(* Logix 5000 project; controller SmartManufacturingCell Emulate 5570 rev 33.11; software revision 33.03; part 2 of 5 *)
(* tags used below, declared in another part *)
   ExitDischargeTimeout : TIMER;   // Non-retentive timer; preset in milliseconds.
   ExitResetONS : BOOL;
   Inspection_RejectSample : BOOL;
   Inspection_StateAtScan : DINT;
   InspectionProcessDelay : TIMER;   // Non-retentive timer; preset in milliseconds.
   InspectionResetONS : BOOL;
   InspectionTimeout : TIMER;   // Non-retentive timer; preset in milliseconds.
   Reject_AutoExtendAllowed : BOOL;
   Reject_ManualExtendAllowed : BOOL;
   Reject_ManualExtendArmed : BOOL;
   Reject_ResetAllowed : BOOL;   // Reject recovery conditions satisfied; permits a fresh Reset request.
   RejectExtendTimeout : TIMER;   // Non-retentive timer; preset in milliseconds.
   RejectResetONS : BOOL;
   RejectRetractTimeout : TIMER;   // Non-retentive timer; preset in milliseconds.
   Cfg_InspectionTimeMs : DINT;   // Inspection duration; 100..2000 ms. Sampled when inspection starts.
   Exit_Flt_DischargeTimeout : BOOL;   // Good or reject bottle departure not confirmed within 3 s Latched; clear cell, remove cause, then fresh Reset.
   Exit_Sts_ResetAccepted : BOOL;   // Exit Sts ResetAccepted
   Exit_Sts_State : DINT;   // 0 Empty; 10 Waiting; 20 Good discharge; 30 Extending; 40 Reject discharge; 50 Retracting; 60 Complete; 90 Faulted
   HMI_Cmd_ClearCell : BOOL;   // Request removal of simulated bottles during fault recovery
   HMI_Cmd_LoadBottle : BOOL;   // Request one simulated bottle at the available entry position
   HMI_Cmd_RejectExtend : BOOL;
   HMI_Cmd_Reset : BOOL;   // Request fault reset after recovery conditions are satisfied
   HMI_Cmd_Stop : BOOL;   // Request controlled production stop
   HMI_Sim_InspectionFailToComplete : BOOL;   // Prevent inspection process timer from completing. Simulation test only.
   HMI_Sim_NextInspectionRejects : BOOL;   // Select Reject for the next inspection
   Inspection_Flt_Timeout : BOOL;   // Inspection did not finish within 3 s Latched; clear cell, remove cause, then fresh Reset.
   Inspection_Sts_ResetAccepted : BOOL;   // Inspection Sts ResetAccepted
   Inspection_Sts_State : DINT;   // 0 Empty; 10 Waiting; 20 Inspecting; 40 Complete; 90 Faulted
   Production_Bottles : UDT_Bottle[4];
   Production_Sts_ClearCellAccepted : BOOL;
   Production_Sts_LoadAccepted : BOOL;
   Production_Sts_LoadAllowed : BOOL;
   Production_Sts_LoadBlockReason : DINT;   // 0 allowed; 10 not Auto Running/ProcessStations; 20 command conflict; 30 conveyor moving; 40 Entry occupied; 50 fault/sta
   Production_Sts_SequenceState : DINT;   // 0 = Idle 10 = ProcessStations 20 = Indexing 30 = ConfirmPositions
   Reject_Flt_FailToExtend : BOOL;   // Reject actuator did not extend within 2 s Latched; clear cell, remove cause, then fresh Reset.
   Reject_Flt_FailToRetract : BOOL;   // Reject actuator did not retract within 2 s Latched; clear cell, remove cause, then fresh Reset.
   Reject_Sts_BlockReason : DINT;   // Reason manual reject extension is unavailable. 0 = Ready to accept Extend. 10 = Release Extend to rearm. 20 = Good-bottl
   Reject_Sts_ResetAccepted : BOOL;
   Sim_In_ConveyorRunning : BOOL;   // Simulated conveyor movement feedback
   Sim_In_EntryPE : BOOL;   // Simulated bottle detected at entry
   Sim_In_GoodExitPE : BOOL;   // Bottle detected passing through good discharge path
   Sim_In_InspectionPE : BOOL;   // Simulated bottle detected at inspection position
   Sim_In_RejectExitPE : BOOL;   // Bottle detected passing through reject discharge path
   Sim_In_RejectExtended : BOOL;   // Simulated reject actuator confirmed extended
   Sim_In_RejectRetracted : BOOL;   // Simulated reject actuator confirmed retracted
   Sim_Out_ConveyorRun : BOOL;   // Command simulated conveyor to run
   Sim_Out_GoodDischargeRun : BOOL;   // Command simulated good-bottle discharge mechanism to run
   Sim_Out_RejectExtend : BOOL;   // Command simulated reject actuator to extend
   Sys_Sts_AutoMode : BOOL;   // Auto mode accepted and active
   Sys_Sts_BlockingFault : BOOL;   // Active blocking fault prevents production and manual equipment operation.
   Sys_Sts_MachineState : DINT;   // 0 = Stopped 10 = Running 20 = Stopping 30 = Faulted
   Sys_Sts_ManualMode : BOOL;   // Manual mode accepted and active
   Sys_Sts_ResetAllowed : BOOL;   // Sys Sts ResetAllowed
   Sys_Sts_StartupReady : BOOL;   // Sys Sts StartupReady
(* Program_Inspection, continued *)

ROUTINE Exit_Faults   (* ladder *)
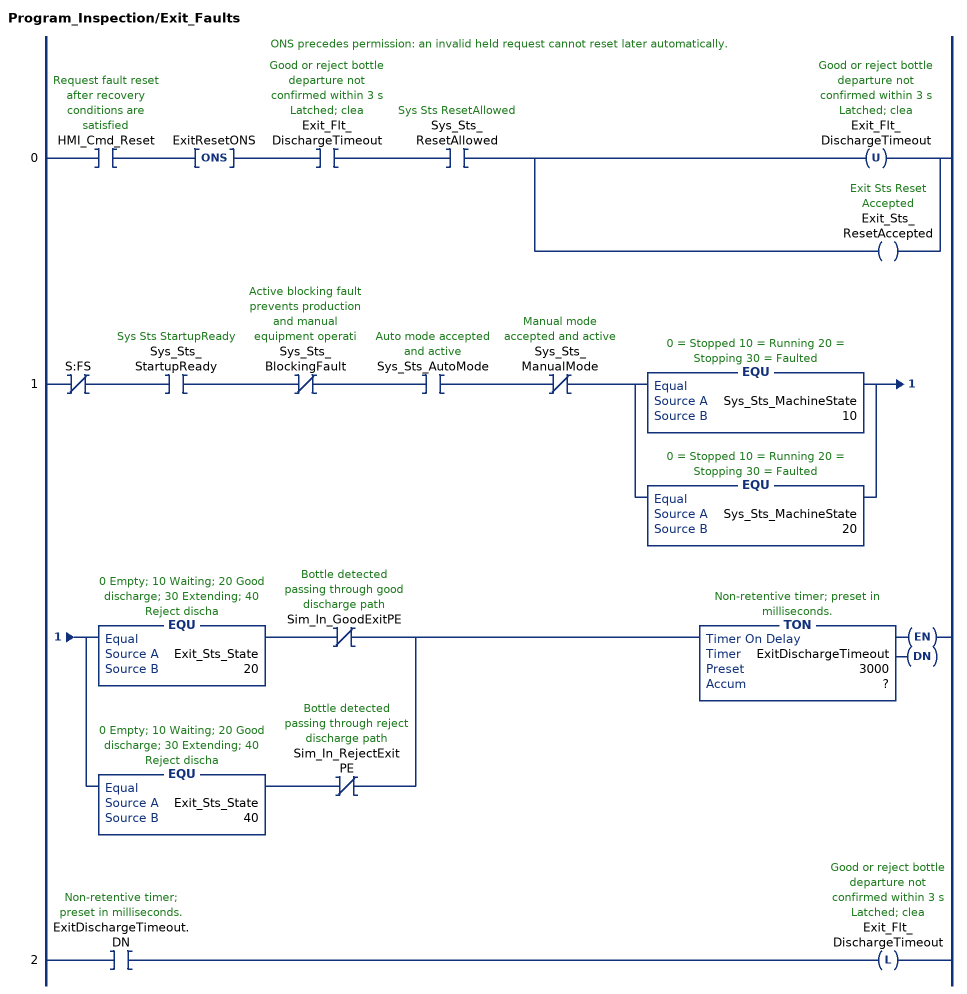
   // ONS precedes permission: an invalid held request cannot reset later automatically.
   0: XIC(HMI_Cmd_Reset)ONS(ExitResetONS)XIC(Exit_Flt_DischargeTimeout)XIC(Sys_Sts_ResetAllowed)[OTU(Exit_Flt_DischargeTimeout) ,OTE(Exit_Sts_ResetAccepted) ];
   1: XIO(S:FS)XIC(Sys_Sts_StartupReady)XIO(Sys_Sts_BlockingFault)XIC(Sys_Sts_AutoMode)XIO(Sys_Sts_ManualMode)[EQU(Sys_Sts_MachineState,10) ,EQU(Sys_Sts_MachineState,20) ][EQU(Exit_Sts_State,20) XIO(Sim_In_GoodExitPE) ,EQU(Exit_Sts_State,40) XIO(Sim_In_RejectExitPE) ]TON(ExitDischargeTimeout,?,?);
   2: XIC(ExitDischargeTimeout.DN)OTL(Exit_Flt_DischargeTimeout);
END_ROUTINE

ROUTINE Inspection_Control   (* ladder *)
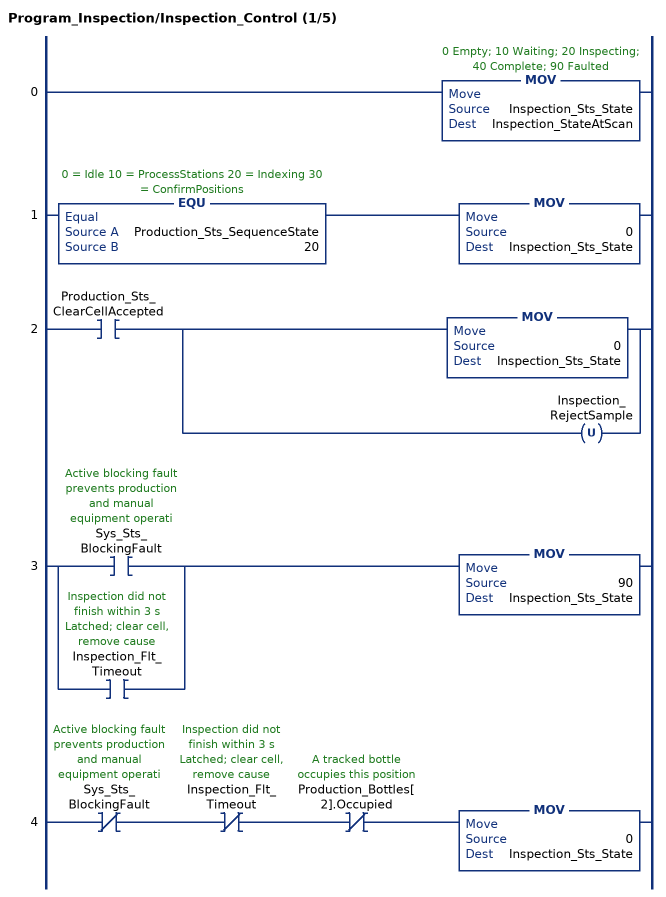
   0: MOV(Inspection_Sts_State,Inspection_StateAtScan);
   1: EQU(Production_Sts_SequenceState,20)MOV(0,Inspection_Sts_State);
   2: XIC(Production_Sts_ClearCellAccepted)[MOV(0,Inspection_Sts_State) ,OTU(Inspection_RejectSample) ];
   3: [XIC(Sys_Sts_BlockingFault) ,XIC(Inspection_Flt_Timeout) ]MOV(90,Inspection_Sts_State);
   4: XIO(Sys_Sts_BlockingFault)XIO(Inspection_Flt_Timeout)XIO(Production_Bottles[2].Occupied)MOV(0,Inspection_Sts_State);
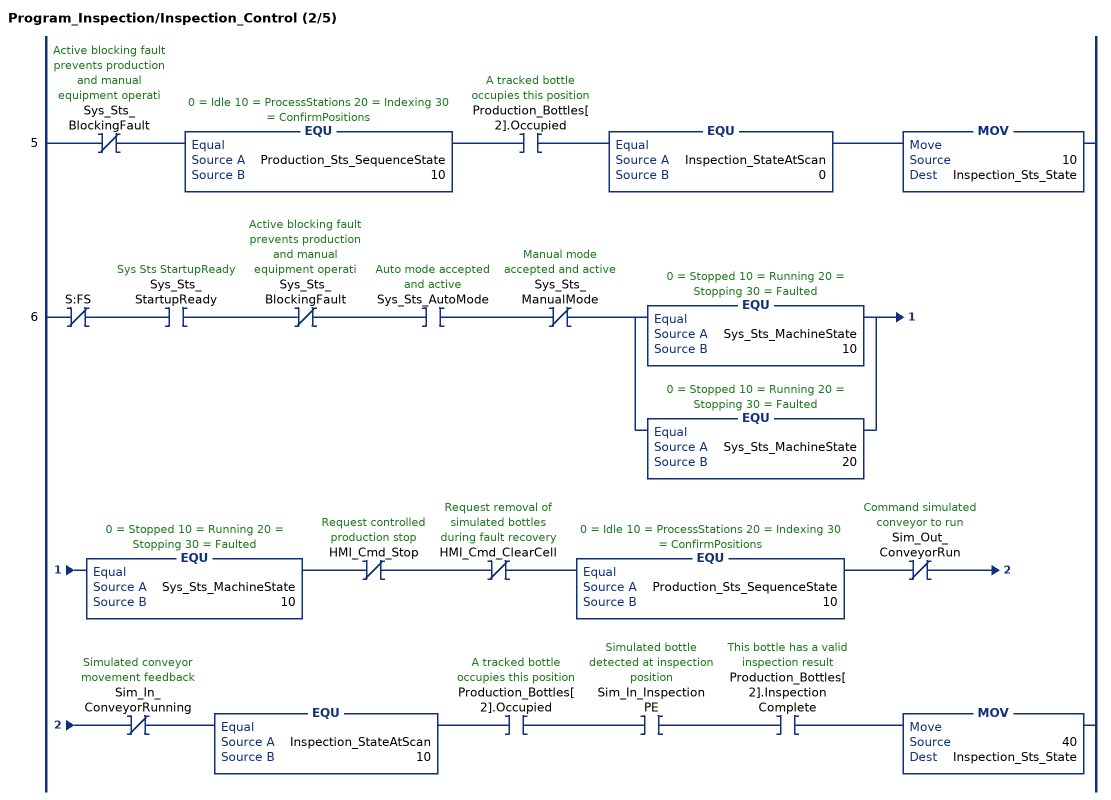
   5: XIO(Sys_Sts_BlockingFault)EQU(Production_Sts_SequenceState,10)XIC(Production_Bottles[2].Occupied)EQU(Inspection_StateAtScan,0)MOV(10,Inspection_Sts_State);
   6: XIO(S:FS)XIC(Sys_Sts_StartupReady)XIO(Sys_Sts_BlockingFault)XIC(Sys_Sts_AutoMode)XIO(Sys_Sts_ManualMode)[EQU(Sys_Sts_MachineState,10) ,EQU(Sys_Sts_MachineState,20) ]EQU(Sys_Sts_MachineState,10)XIO(HMI_Cmd_Stop)XIO(HMI_Cmd_ClearCell)EQU(Production_Sts_SequenceState,10)XIO(Sim_Out_ConveyorRun)XIO(Sim_In_ConveyorRunning)EQU(Inspection_StateAtScan,10)XIC(Production_Bottles[2].Occupied)XIC(Sim_In_InspectionPE)XIC(Production_Bottles[2].InspectionComplete)MOV(40,Inspection_Sts_State);
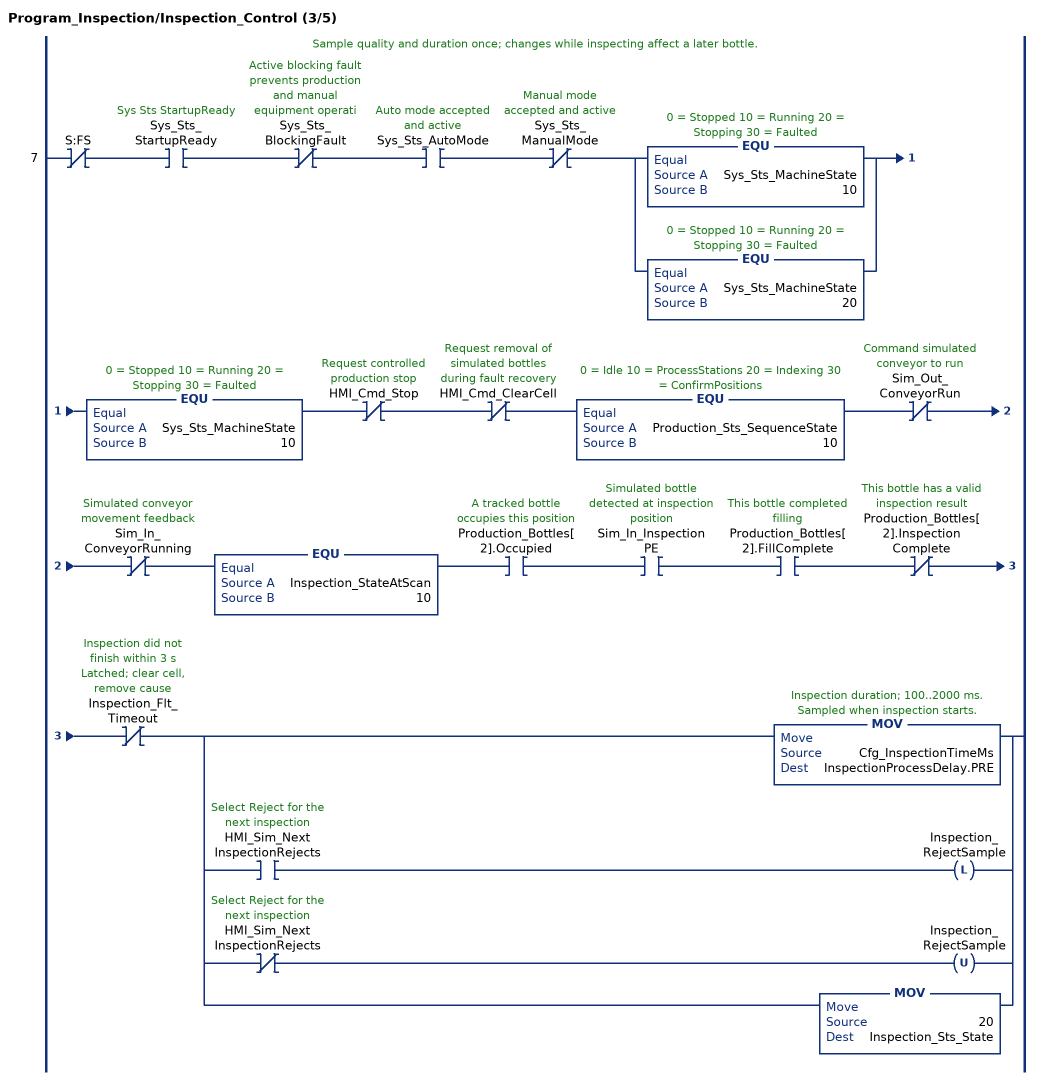
   // Sample quality and duration once; changes while inspecting affect a later bottle.
   7: XIO(S:FS)XIC(Sys_Sts_StartupReady)XIO(Sys_Sts_BlockingFault)XIC(Sys_Sts_AutoMode)XIO(Sys_Sts_ManualMode)[EQU(Sys_Sts_MachineState,10) ,EQU(Sys_Sts_MachineState,20) ]EQU(Sys_Sts_MachineState,10)XIO(HMI_Cmd_Stop)XIO(HMI_Cmd_ClearCell)EQU(Production_Sts_SequenceState,10)XIO(Sim_Out_ConveyorRun)XIO(Sim_In_ConveyorRunning)EQU(Inspection_StateAtScan,10)XIC(Production_Bottles[2].Occupied)XIC(Sim_In_InspectionPE)XIC(Production_Bottles[2].FillComplete)XIO(Production_Bottles[2].InspectionComplete)XIO(Inspection_Flt_Timeout)[MOV(Cfg_InspectionTimeMs,InspectionProcessDelay.PRE) ,XIC(HMI_Sim_NextInspectionRejects) OTL(Inspection_RejectSample) ,XIO(HMI_Sim_NextInspectionRejects) OTU(Inspection_RejectSample) ,MOV(20,Inspection_Sts_State) ];
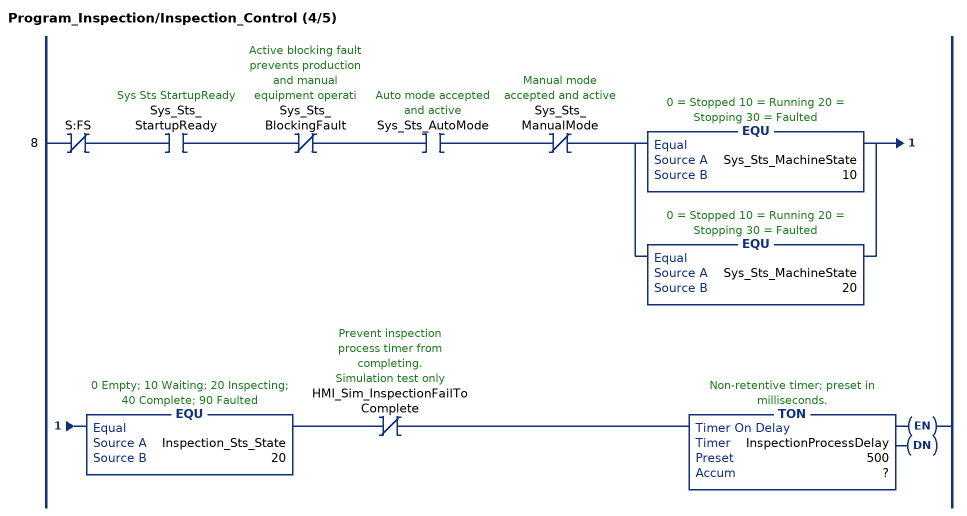
   8: XIO(S:FS)XIC(Sys_Sts_StartupReady)XIO(Sys_Sts_BlockingFault)XIC(Sys_Sts_AutoMode)XIO(Sys_Sts_ManualMode)[EQU(Sys_Sts_MachineState,10) ,EQU(Sys_Sts_MachineState,20) ]EQU(Inspection_Sts_State,20)XIO(HMI_Sim_InspectionFailToComplete)TON(InspectionProcessDelay,?,?);
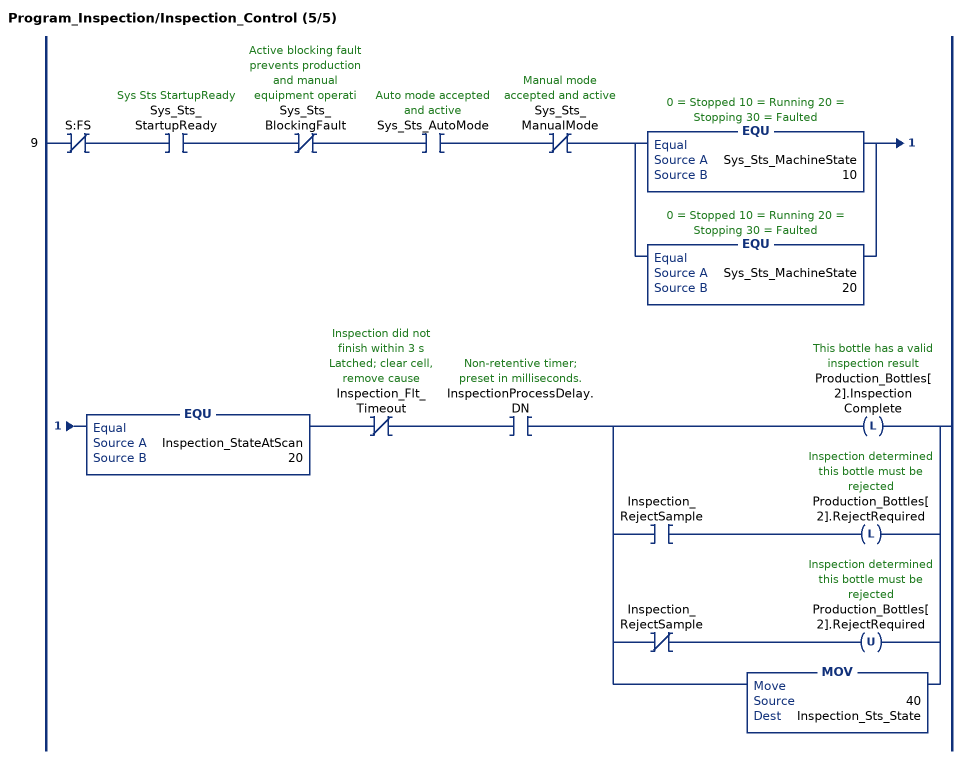
   9: XIO(S:FS)XIC(Sys_Sts_StartupReady)XIO(Sys_Sts_BlockingFault)XIC(Sys_Sts_AutoMode)XIO(Sys_Sts_ManualMode)[EQU(Sys_Sts_MachineState,10) ,EQU(Sys_Sts_MachineState,20) ]EQU(Inspection_StateAtScan,20)XIO(Inspection_Flt_Timeout)XIC(InspectionProcessDelay.DN)[OTL(Production_Bottles[2].InspectionComplete) ,XIC(Inspection_RejectSample) OTL(Production_Bottles[2].RejectRequired) ,XIO(Inspection_RejectSample) OTU(Production_Bottles[2].RejectRequired) ,MOV(40,Inspection_Sts_State) ];
END_ROUTINE

ROUTINE Inspection_Faults   (* ladder *)
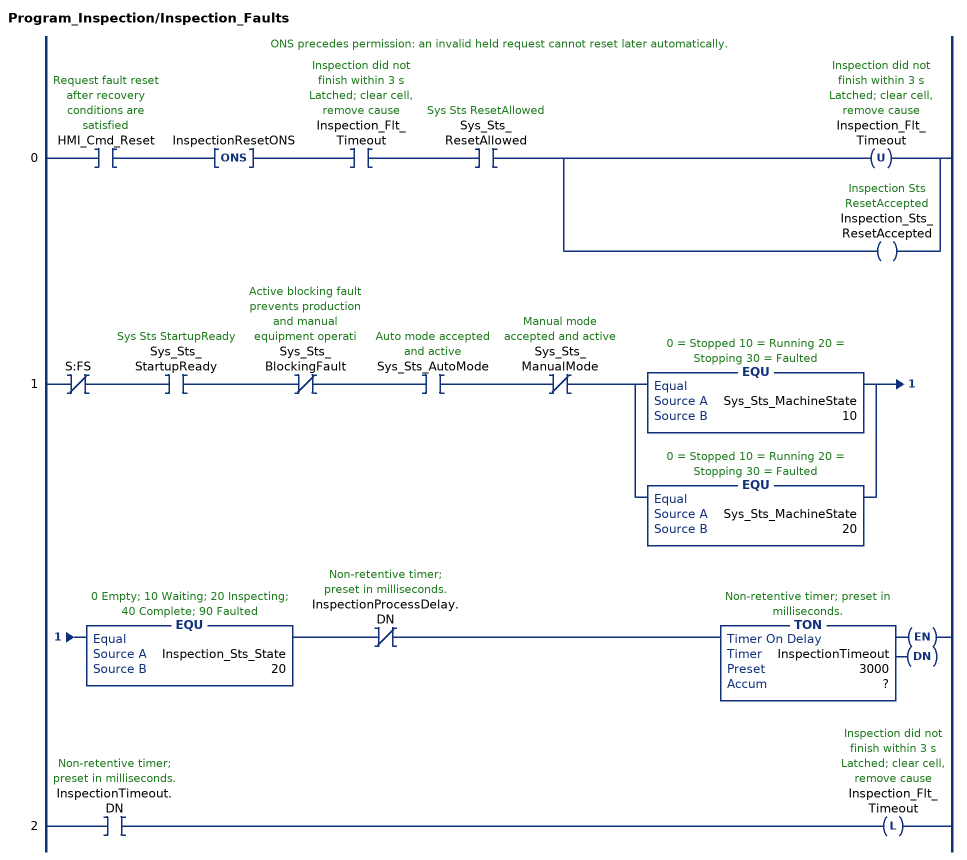
   // ONS precedes permission: an invalid held request cannot reset later automatically.
   0: XIC(HMI_Cmd_Reset)ONS(InspectionResetONS)XIC(Inspection_Flt_Timeout)XIC(Sys_Sts_ResetAllowed)[OTU(Inspection_Flt_Timeout) ,OTE(Inspection_Sts_ResetAccepted) ];
   1: XIO(S:FS)XIC(Sys_Sts_StartupReady)XIO(Sys_Sts_BlockingFault)XIC(Sys_Sts_AutoMode)XIO(Sys_Sts_ManualMode)[EQU(Sys_Sts_MachineState,10) ,EQU(Sys_Sts_MachineState,20) ]EQU(Inspection_Sts_State,20)XIO(InspectionProcessDelay.DN)TON(InspectionTimeout,?,?);
   2: XIC(InspectionTimeout.DN)OTL(Inspection_Flt_Timeout);
END_ROUTINE

ROUTINE MainRoutine   (* ladder *)
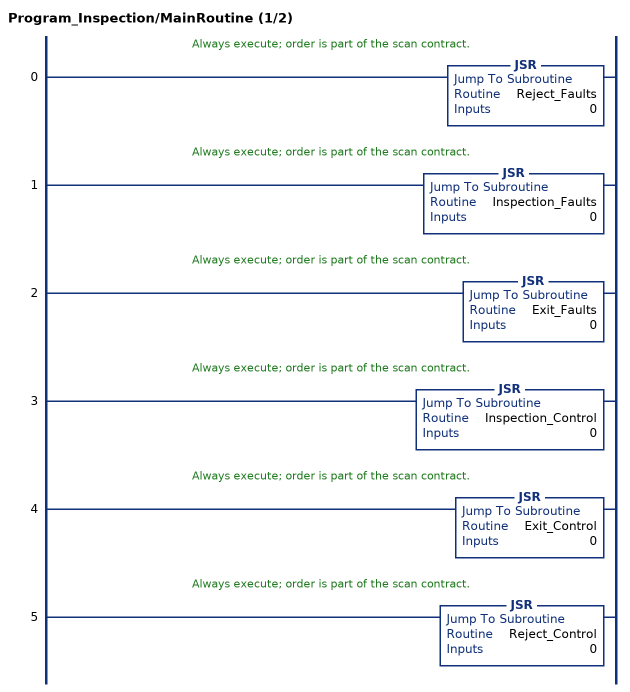
   // Always execute; order is part of the scan contract.
   0: JSR(Reject_Faults,0);
   // Always execute; order is part of the scan contract.
   1: JSR(Inspection_Faults,0);
   // Always execute; order is part of the scan contract.
   2: JSR(Exit_Faults,0);
   // Always execute; order is part of the scan contract.
   3: JSR(Inspection_Control,0);
   // Always execute; order is part of the scan contract.
   4: JSR(Exit_Control,0);
   // Always execute; order is part of the scan contract.
   5: JSR(Reject_Control,0);
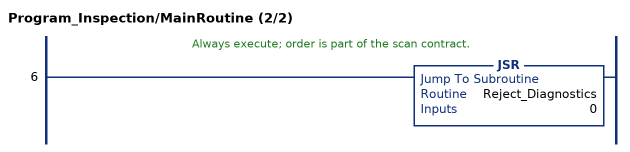
   // Always execute; order is part of the scan contract.
   6: JSR(Reject_Diagnostics,0);
END_ROUTINE

ROUTINE Reject_Control   (* ladder *)
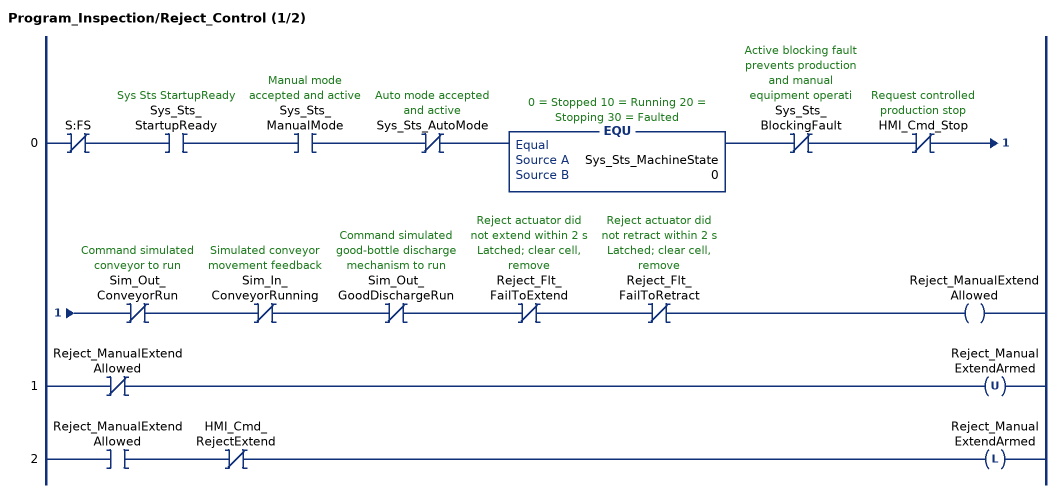
   0: XIO(S:FS)XIC(Sys_Sts_StartupReady)XIC(Sys_Sts_ManualMode)XIO(Sys_Sts_AutoMode)EQU(Sys_Sts_MachineState,0)XIO(Sys_Sts_BlockingFault)XIO(HMI_Cmd_Stop)XIO(Sim_Out_ConveyorRun)XIO(Sim_In_ConveyorRunning)XIO(Sim_Out_GoodDischargeRun)XIO(Reject_Flt_FailToExtend)XIO(Reject_Flt_FailToRetract)OTE(Reject_ManualExtendAllowed);
   1: XIO(Reject_ManualExtendAllowed)OTU(Reject_ManualExtendArmed);
   2: XIC(Reject_ManualExtendAllowed)XIO(HMI_Cmd_RejectExtend)OTL(Reject_ManualExtendArmed);
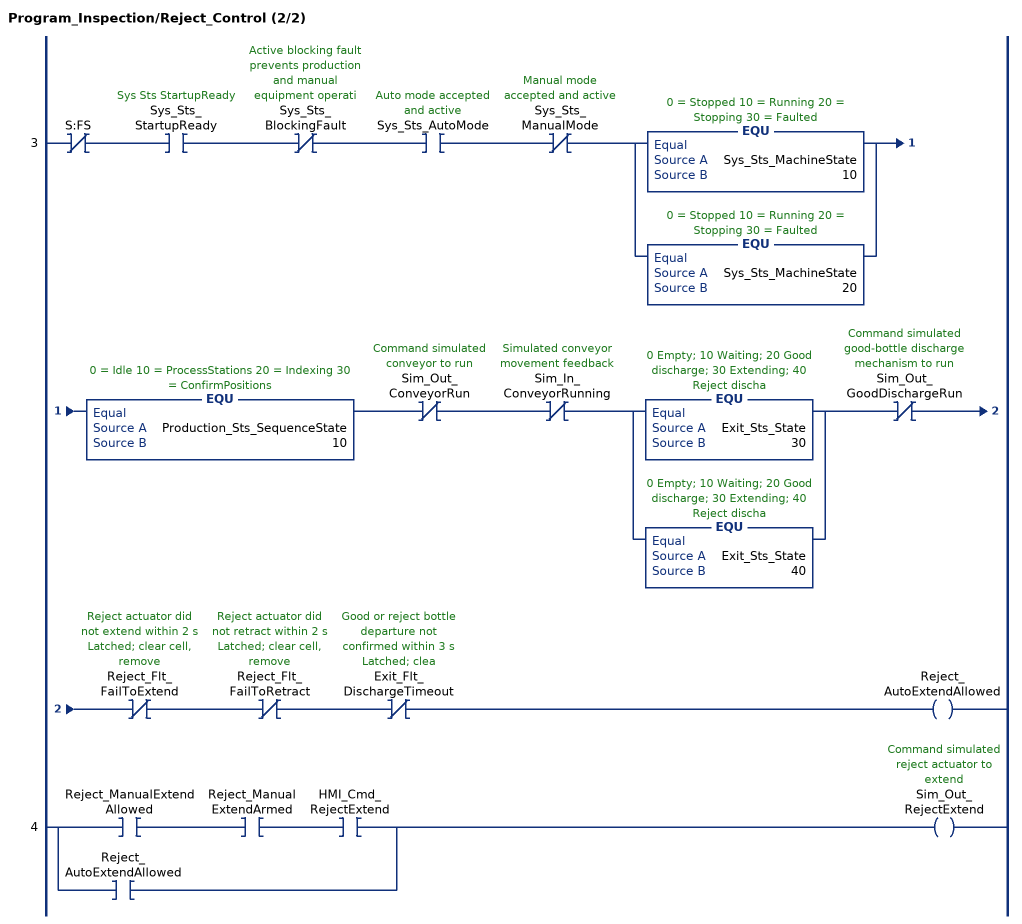
   3: XIO(S:FS)XIC(Sys_Sts_StartupReady)XIO(Sys_Sts_BlockingFault)XIC(Sys_Sts_AutoMode)XIO(Sys_Sts_ManualMode)[EQU(Sys_Sts_MachineState,10) ,EQU(Sys_Sts_MachineState,20) ]EQU(Production_Sts_SequenceState,10)XIO(Sim_Out_ConveyorRun)XIO(Sim_In_ConveyorRunning)[EQU(Exit_Sts_State,30) ,EQU(Exit_Sts_State,40) ]XIO(Sim_Out_GoodDischargeRun)XIO(Reject_Flt_FailToExtend)XIO(Reject_Flt_FailToRetract)XIO(Exit_Flt_DischargeTimeout)OTE(Reject_AutoExtendAllowed);
   4: [XIC(Reject_ManualExtendAllowed) XIC(Reject_ManualExtendArmed) XIC(HMI_Cmd_RejectExtend) ,XIC(Reject_AutoExtendAllowed) ]OTE(Sim_Out_RejectExtend);
END_ROUTINE

ROUTINE Reject_Diagnostics   (* ladder *)
// Reason manual reject extension is unavailable
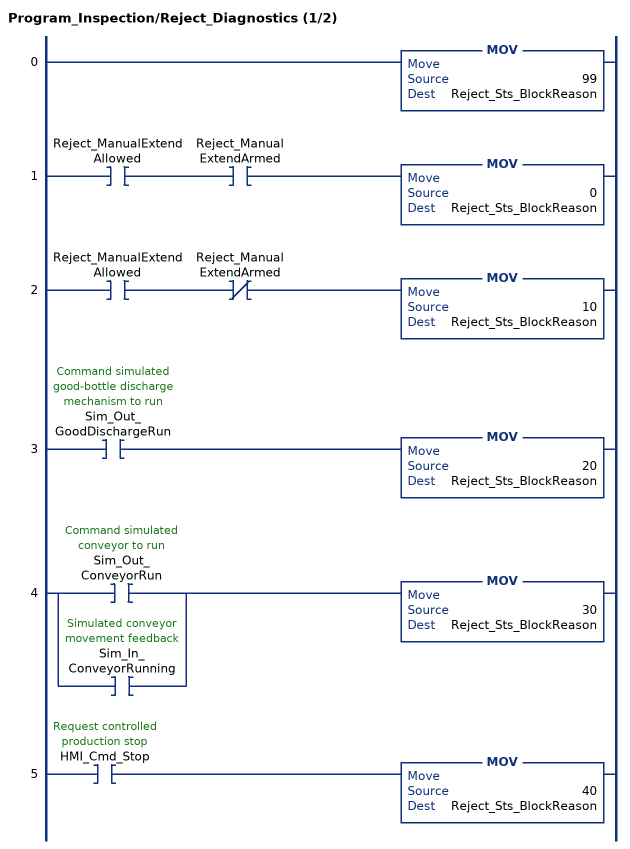
   0: MOV(99,Reject_Sts_BlockReason);
   1: XIC(Reject_ManualExtendAllowed)XIC(Reject_ManualExtendArmed)MOV(0,Reject_Sts_BlockReason);
   2: XIC(Reject_ManualExtendAllowed)XIO(Reject_ManualExtendArmed)MOV(10,Reject_Sts_BlockReason);
   3: XIC(Sim_Out_GoodDischargeRun)MOV(20,Reject_Sts_BlockReason);
   4: [XIC(Sim_Out_ConveyorRun) ,XIC(Sim_In_ConveyorRunning) ]MOV(30,Reject_Sts_BlockReason);
   5: XIC(HMI_Cmd_Stop)MOV(40,Reject_Sts_BlockReason);
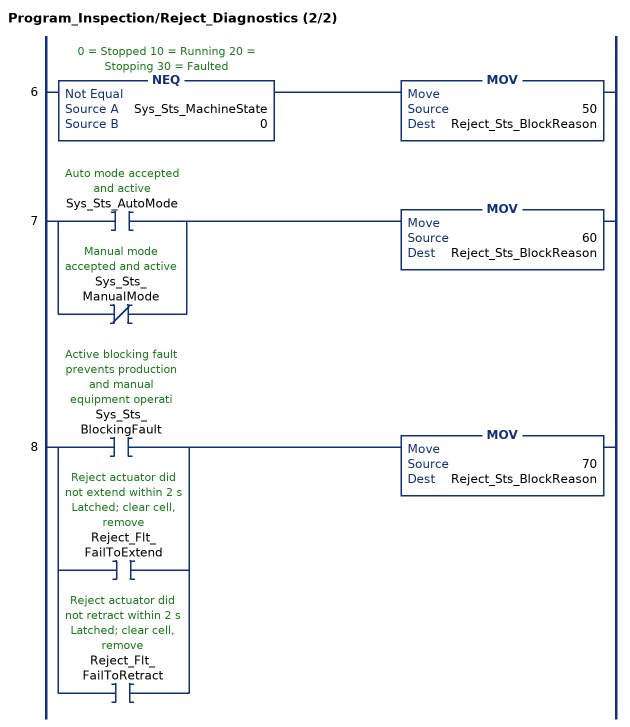
   6: NEQ(Sys_Sts_MachineState,0)MOV(50,Reject_Sts_BlockReason);
   7: [XIC(Sys_Sts_AutoMode) ,XIO(Sys_Sts_ManualMode) ]MOV(60,Reject_Sts_BlockReason);
   8: [XIC(Sys_Sts_BlockingFault) ,XIC(Reject_Flt_FailToExtend) ,XIC(Reject_Flt_FailToRetract) ]MOV(70,Reject_Sts_BlockReason);
END_ROUTINE

ROUTINE Reject_Faults   (* ladder *)
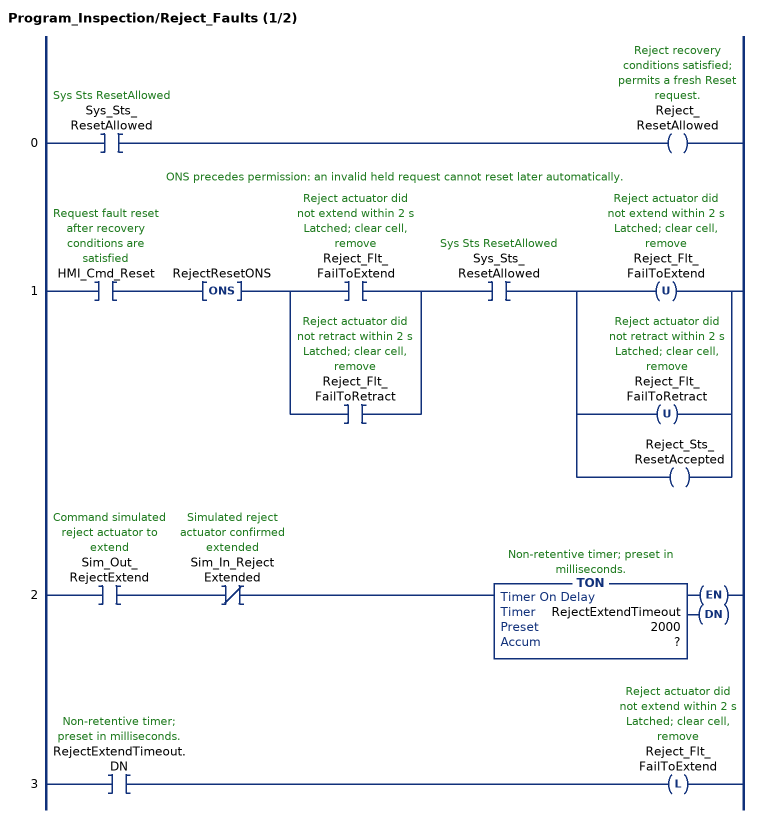
   0: XIC(Sys_Sts_ResetAllowed)OTE(Reject_ResetAllowed);
   // ONS precedes permission: an invalid held request cannot reset later automatically.
   1: XIC(HMI_Cmd_Reset)ONS(RejectResetONS)[XIC(Reject_Flt_FailToExtend) ,XIC(Reject_Flt_FailToRetract) ]XIC(Sys_Sts_ResetAllowed)[OTU(Reject_Flt_FailToExtend) ,OTU(Reject_Flt_FailToRetract) ,OTE(Reject_Sts_ResetAccepted) ];
   2: XIC(Sim_Out_RejectExtend)XIO(Sim_In_RejectExtended)TON(RejectExtendTimeout,?,?);
   3: XIC(RejectExtendTimeout.DN)OTL(Reject_Flt_FailToExtend);
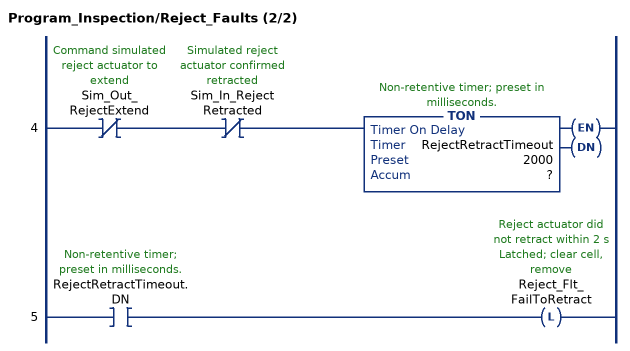
   4: XIO(Sim_Out_RejectExtend)XIO(Sim_In_RejectRetracted)TON(RejectRetractTimeout,?,?);
   5: XIC(RejectRetractTimeout.DN)OTL(Reject_Flt_FailToRetract);
END_ROUTINE
END_PROGRAM

PROGRAM Program_Production   (* main routine MainRoutine *)
// Production sequence coordination, bottle tracking, and production statistics.
VAR
   ClearCell_CommandsReleased : BOOL; {access None}
   ClearCell_EquipmentReady : BOOL; {access None}
   ClearCellRequestONS : BOOL; {access None}
   Exit_ReadyForIndex : BOOL; {access None}
   Filling_ReadyForIndex : BOOL; {access None}
   Index_CommandsReleased : BOOL; {access None}
   Index_EquipmentReady : BOOL; {access None}
   IndexConfirmTimeout : TIMER := (PRE := 1000); {access None}   // Non-retentive timer; preset in milliseconds.
   IndexTimeout : TIMER := (PRE := 3000); {access None}   // Non-retentive timer; preset in milliseconds.
   Inspection_ReadyForIndex : BOOL; {access None}
   LoadRequestONS : BOOL; {access None}
   Production_CycleHealthy : BOOL; {access None}
   Production_ResetAllowed : BOOL; {access None}
   Production_ResetCommandsReleased : BOOL; {access None}
   Production_SensorsClear : BOOL; {access None}
   Production_TrackingEmpty : BOOL; {access None}
   ProductionResetONS : BOOL; {access None}
   SequenceAtScan : DINT; {access None}
   StatisticsResetAccepted : BOOL; {access None}
   StatisticsResetONS : BOOL; {access None}
   Stats_ExitElapsed : REAL; {access None}
   Stats_HasPreviousExit : BOOL; {access None}
   Stats_RateElapsed : REAL; {access None}
   Stats_WindowCount : DINT; {access None}
   TrackingMismatchDelay : TIMER := (PRE := 200); {access None}   // Non-retentive timer; preset in milliseconds.
END_VAR

ROUTINE Bottle_Loading   (* ladder *)
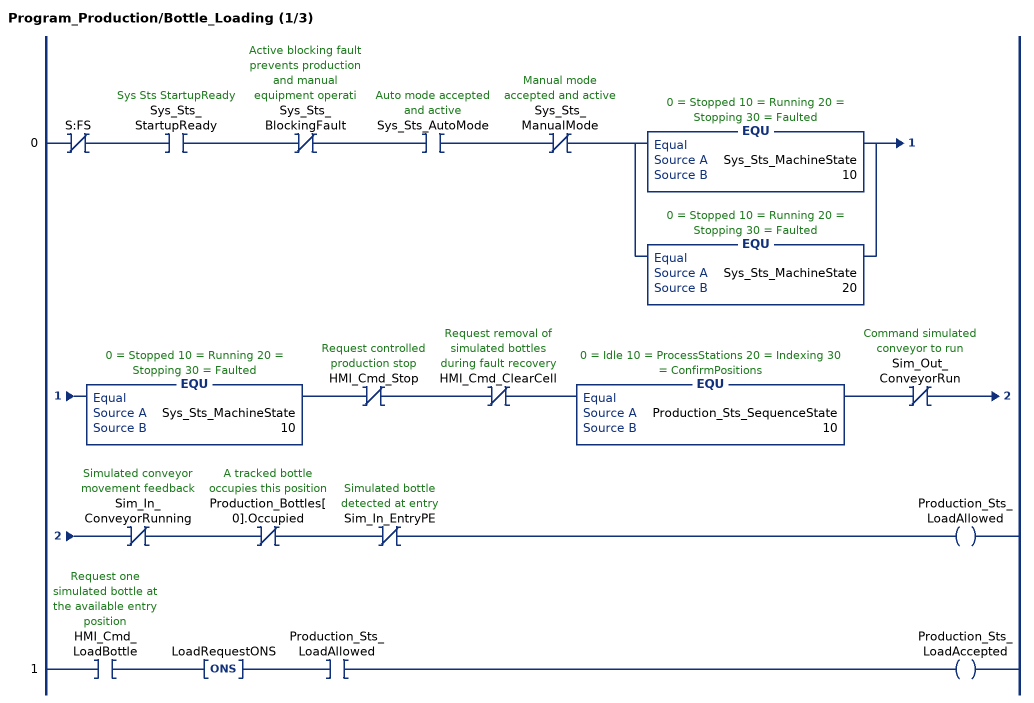
   0: XIO(S:FS)XIC(Sys_Sts_StartupReady)XIO(Sys_Sts_BlockingFault)XIC(Sys_Sts_AutoMode)XIO(Sys_Sts_ManualMode)[EQU(Sys_Sts_MachineState,10) ,EQU(Sys_Sts_MachineState,20) ]EQU(Sys_Sts_MachineState,10)XIO(HMI_Cmd_Stop)XIO(HMI_Cmd_ClearCell)EQU(Production_Sts_SequenceState,10)XIO(Sim_Out_ConveyorRun)XIO(Sim_In_ConveyorRunning)XIO(Production_Bottles[0].Occupied)XIO(Sim_In_EntryPE)OTE(Production_Sts_LoadAllowed);
   1: XIC(HMI_Cmd_LoadBottle)ONS(LoadRequestONS)XIC(Production_Sts_LoadAllowed)OTE(Production_Sts_LoadAccepted);
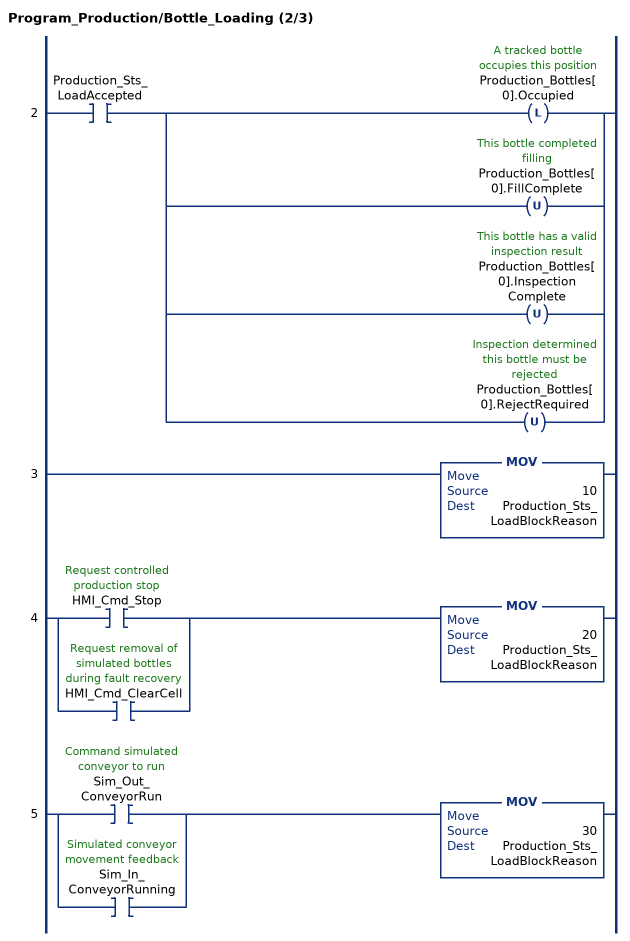
   2: XIC(Production_Sts_LoadAccepted)[OTL(Production_Bottles[0].Occupied) ,OTU(Production_Bottles[0].FillComplete) ,OTU(Production_Bottles[0].InspectionComplete) ,OTU(Production_Bottles[0].RejectRequired) ];
   3: MOV(10,Production_Sts_LoadBlockReason);
   4: [XIC(HMI_Cmd_Stop) ,XIC(HMI_Cmd_ClearCell) ]MOV(20,Production_Sts_LoadBlockReason);
   5: [XIC(Sim_Out_ConveyorRun) ,XIC(Sim_In_ConveyorRunning) ]MOV(30,Production_Sts_LoadBlockReason);
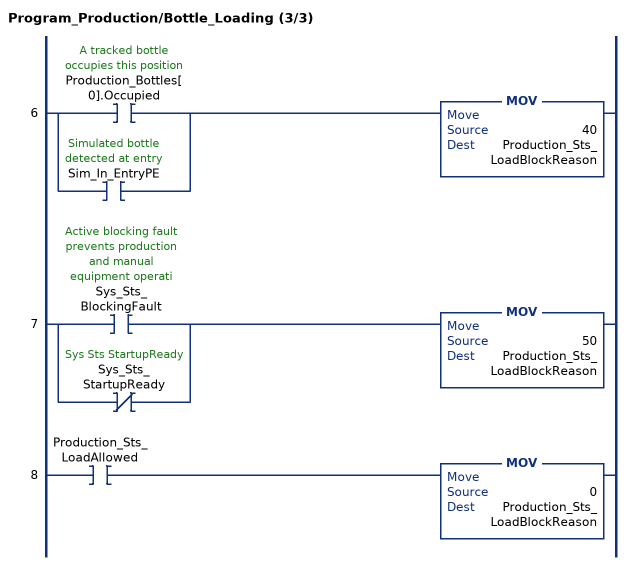
   6: [XIC(Production_Bottles[0].Occupied) ,XIC(Sim_In_EntryPE) ]MOV(40,Production_Sts_LoadBlockReason);
   7: [XIC(Sys_Sts_BlockingFault) ,XIO(Sys_Sts_StartupReady) ]MOV(50,Production_Sts_LoadBlockReason);
   8: XIC(Production_Sts_LoadAllowed)MOV(0,Production_Sts_LoadBlockReason);
END_ROUTINE
